Fanuc KAREL source: kt00033.KL

PROGRAM KT00033
%NOLOCKGROUP
VAR
I1:INTEGER;I2:INTEGER;OUT:INTEGER
BEGIN
--
--
I1=2
I2=3
I1=2
I2=3
OUT=(I1-I2)
END KT00033
